TYPE "ST_PartResult"
VERSION : 0.1
   STRUCT
      Verdict : DInt;
      ReasonCode : DInt;
      Records : Array[1..32] of "ST_MeasRecord";
      StationPath : WString[255];
      Stamp : LDT;
      TimeSynchronized : Bool;
   END_STRUCT;

END_TYPE

